TYPE "FRK_Document_D012"
VERSION : 0.1
   STRUCT
      "SchemaVersion" {ExternalAccessible := 'False'; ExternalVisible := 'False'; ExternalWritable := 'False'} : UInt;
      "Scope" {ExternalAccessible := 'False'; ExternalVisible := 'False'; ExternalWritable := 'False'} : String[80];
      "Image" {ExternalAccessible := 'False'; ExternalVisible := 'False'; ExternalWritable := 'False'} : "FRK_ModelImage";
   END_STRUCT;
END_TYPE
